(* PLC project ExampleProject, Example Org Example IDE 1.0 *)
(* stored: creationDateTime 2026-01-05T08:00:00, version 1, modificationDateTime 2026-11-01T03:12:00 *)

TYPE ST_ExamplePump : STRUCT
  SpeedSP : REAL := 0.0;
  FaultCode : DINT;
END_STRUCT;
END_TYPE

FUNCTION_BLOCK FB_ExampleValve
  VAR_INPUT
    OpenCmd : BOOL;
    Permissive : BOOL;
    Bypass : BOOL;
  END_VAR
  VAR_OUTPUT
    OpenOut : BOOL;
  END_VAR

OpenOut := OpenCmd OR Bypass; (* permissive required *)
END_FUNCTION_BLOCK

PROGRAM PLC_PRG
  VAR
    Run : BOOL;  (* Example run command from the HMI *)
    Pump1 : ST_ExamplePump;
    Valve1 : FB_ExampleValve;
  END_VAR
  VAR CONSTANT
    HighLimit : REAL := 95.0;
  END_VAR

// Example speed clamp
IF Pump1.SpeedSP > HighLimit THEN
    Pump1.SpeedSP := HighLimit + 20.0;
END_IF;
Valve1(OpenCmd := Run, Permissive := Pump1.SpeedSP < HighLimit);
END_PROGRAM

CONFIGURATION ExampleConfig
  RESOURCE ExampleResource ON PLC
    TASK MainTask(INTERVAL := T#100ms, PRIORITY := 1);
    PROGRAM PLC_PRG WITH MainTask : PLC_PRG;
  END_RESOURCE
END_CONFIGURATION
